{attribute 'no_explicit_call':= 'do not call this POU directly'}
FUNCTION_BLOCK T_DetectOnlineChange
VAR
    StoredOnlineChangeCnt : UDINT := 99;
	_OnlineChangeDetected : BOOL;
END_VAR

METHOD CyclicUpdate
IF TwinCAT_SystemInfoVarList._AppInfo.OnlineChangeCnt <> StoredOnlineChangeCnt THEN
    _OnlineChangeDetected  := TRUE;
    StoredOnlineChangeCnt := TwinCAT_SystemInfoVarList._AppInfo.OnlineChangeCnt;
END_IF
END_METHOD

PROPERTY OnlineChangeDetected : BOOL
GET
OnlineChangeDetected := _OnlineChangeDetected;
END_GET
END_PROPERTY

END_FUNCTION_BLOCK

(* stored: Version 1.1.0.1, ProductVersion 3.1.4026.19
   POU T_DetectOnlineChange: Id {424d8bc0-80ad-4ff2-af04-d54ec3aa7c3d}, SpecialFunc None
   Method CyclicUpdate: Id {ca6150a4-825e-4ae2-a66d-4ccf39e851c0}
   Property OnlineChangeDetected: Id {8b032061-7ebc-4bef-90b5-0185eb36d1fc}
   Get Get: Id {fe7cfc2e-5c73-4d4f-b1ce-90d3f01b68df} *)
